(* IEC 61131-3 sources: plc-vscode/tests/st/test-ready/rusty/tests/lit/single/conversion, 6 files *)

(* ---- real_trunc_int.st ---- *)
// RUN: (%COMPILE %s && %RUN) | %CHECK %s
FUNCTION main
    printf('%d$N', REAL_TRUNC_SINT(5.6));       // CHECK: 5
    printf('%d$N', REAL_TRUNC_USINT(5.6));      // CHECK: 5
    printf('%d$N', REAL_TRUNC_INT(5.6));        // CHECK: 5
    printf('%d$N', REAL_TRUNC_UINT(5.6));       // CHECK: 5
    printf('%d$N', REAL_TRUNC_INT(5.6));        // CHECK: 5
    printf('%d$N', REAL_TRUNC_UINT(5.6));       // CHECK: 5
    printf('%d$N', REAL_TRUNC_DINT(5.6));       // CHECK: 5
    printf('%d$N', REAL_TRUNC_UDINT(5.6));      // CHECK: 5
    printf('%d$N', REAL_TRUNC_LINT(5.6));       // CHECK: 5
    printf('%d$N', REAL_TRUNC_ULINT(5.6));      // CHECK: 5

    printf('%d$N', REAL_TRUNC_SINT(-5.6));      // CHECK: -5
    printf('%d$N', REAL_TRUNC_INT(-5.6));       // CHECK: -5
    printf('%d$N', REAL_TRUNC_DINT(-5.6));      // CHECK: -5
    printf('%d$N', REAL_TRUNC_LINT(-5.6));      // CHECK: -5
END_FUNCTION

(* ---- to_bit.st ---- *)
// Note: Tests are kept simple because there are already tests covering the underliny X_TO_Y functions, which
//       the TO_Y(X) functions are based on.

// RUN: (%COMPILE %s && %RUN) | %CHECK %s
FUNCTION main
    printf('%d$N', TO_BOOL(BOOL#FALSE));        // CHECK: 0
    printf('%d$N', TO_BOOL(BOOL#TRUE));         // CHECK: 1
    printf('%d$N', TO_BOOL(BYTE#0));            // CHECK: 0
    printf('%d$N', TO_BOOL(BYTE#5));            // CHECK: 1
    printf('%d$N', TO_BOOL(WORD#0));            // CHECK: 0
    printf('%d$N', TO_BOOL(WORD#5));            // CHECK: 1
    printf('%d$N', TO_BOOL(DWORD#0));           // CHECK: 0
    printf('%d$N', TO_BOOL(DWORD#5));           // CHECK: 1
    printf('%d$N', TO_BOOL(LWORD#0));           // CHECK: 0
    printf('%d$N', TO_BOOL(LWORD#5));           // CHECK: 1

    printf('%d$N', TO_BYTE(BYTE#5));            // CHECK: 5
    printf('%d$N', TO_BYTE(BOOL#FALSE));        // CHECK: 0
    printf('%d$N', TO_BYTE(BOOL#TRUE));         // CHECK: 1
    printf('%d$N', TO_BYTE(CHAR#'a'));          // CHECK: 97
    printf('%d$N', TO_BYTE(WCHAR#"a"));         // CHECK: 97
    printf('%d$N', TO_BYTE(WORD#5));            // CHECK: 5
    printf('%d$N', TO_BYTE(DWORD#5));           // CHECK: 5
    printf('%d$N', TO_BYTE(LWORD#5));           // CHECK: 5

    printf('%d$N', TO_WORD(WORD#5));            // CHECK: 5
    printf('%d$N', TO_WORD(BOOL#FALSE));        // CHECK: 0
    printf('%d$N', TO_WORD(BOOL#TRUE));         // CHECK: 1
    printf('%d$N', TO_WORD(CHAR#'a'));          // CHECK: 97
    printf('%d$N', TO_WORD(WCHAR#"a"));         // CHECK: 97
    printf('%d$N', TO_WORD(BYTE#5));            // CHECK: 5
    printf('%d$N', TO_WORD(DWORD#5));           // CHECK: 5
    printf('%d$N', TO_WORD(LWORD#5));           // CHECK: 5

    printf('%d$N', TO_DWORD(DWORD#5));          // CHECK: 5
    printf('%d$N', TO_DWORD(BOOL#FALSE));       // CHECK: 0
    printf('%d$N', TO_DWORD(BOOL#TRUE));        // CHECK: 1
    printf('%d$N', TO_DWORD(CHAR#'a'));         // CHECK: 97
    printf('%d$N', TO_DWORD(WCHAR#'a'));        // CHECK: 97
    printf('%d$N', TO_DWORD(BYTE#5));           // CHECK: 5
    printf('%d$N', TO_DWORD(WORD#5));           // CHECK: 5
    printf('%d$N', TO_DWORD(LWORD#5));          // CHECK: 5

    printf('%d$N', TO_LWORD(LWORD#5));          // CHECK: 5
    printf('%d$N', TO_LWORD(BOOL#FALSE));       // CHECK: 0
    printf('%d$N', TO_LWORD(BOOL#TRUE));        // CHECK: 1
    printf('%d$N', TO_LWORD(CHAR#'a'));         // CHECK: 97
    printf('%d$N', TO_LWORD(WCHAR#'a'));        // CHECK: 97
    printf('%d$N', TO_LWORD(BYTE#5));           // CHECK: 5
    printf('%d$N', TO_LWORD(WORD#5));           // CHECK: 5
    printf('%d$N', TO_LWORD(DWORD#5));          // CHECK: 5
END_FUNCTION

(* ---- to_date_time.st ---- *)
// RUN: (%COMPILE %s && %RUN) | %CHECK %s
FUNCTION main
    // TO_TIME
    printf('%s$N', REF(TIME_TO_STRING(TO_TIME(LTIME#10s))));                        // CHECK: 10s

    // TO_LTIME
    printf('%s$N', REF(TIME_TO_STRING(TO_LTIME(TIME#10s))));                        // CHECK: 10s

    // TO_DT
    printf('%s$N', REF(TIME_TO_STRING(TO_DT(LDT#2024-11-12-16:36:15.100))));        // CHECK: 20039d16h36m15s100ms

    // TO_LDT
    printf('%s$N', REF(TIME_TO_STRING(TO_LDT(DT#2024-11-12-16:36:15.100))));        // CHECK: 20039d16h36m15s100ms

    // TO_DATE
    printf('%s$N', REF(TIME_TO_STRING(TO_DATE(DT#2024-11-12-16:36:15.100))));       // CHECK: 20039d
    printf('%s$N', REF(TIME_TO_STRING(TO_DATE(LDT#2024-11-12-16:36:15.100))));      // CHECK: 20039d

    // TO_LDATE
    printf('%s$N', REF(TIME_TO_STRING(TO_LDATE(DT#2024-11-12-16:36:15.100))));       // CHECK: 20039d
    printf('%s$N', REF(TIME_TO_STRING(TO_LDATE(LDT#2024-11-12-16:36:15.100))));      // CHECK: 20039d

    // TO_TOD
    printf('%s$N', REF(LTOD_TO_STRING(TO_TOD(LTOD#16:36:15))));                     // CHECK: 16:36:15
    printf('%s$N', REF(TOD_TO_STRING(TO_TOD(DT#2024-11-12-16:36:15.100))));         // CHECK: 16:36:15.100
    printf('%s$N', REF(TOD_TO_STRING(TO_TOD(LDT#2024-11-12-16:36:15.100))));        // CHECK: 16:36:15.100

    // TO_LTOD
    printf('%s$N', REF(LTOD_TO_STRING(TO_LTOD(TOD#16:36:15))));                     // CHECK: 16:36:15
    printf('%s$N', REF(LTOD_TO_STRING(TO_LTOD(DT#2024-11-12-16:36:15.100))));       // CHECK: 16:36:15.100
    printf('%s$N', REF(LTOD_TO_STRING(TO_LTOD(LDT#2024-11-12-16:36:15.100))));      // CHECK: 16:36:15.100
END_FUNCTION

(* ---- to_num.st ---- *)
// RUN: (%COMPILE %s && %RUN) | %CHECK %s
FUNCTION main
    printf('%d$N', TO_SINT(SINT#5));            // CHECK: 5
    printf('%d$N', TO_SINT(USINT#5));           // CHECK: 5
    printf('%d$N', TO_SINT(INT#5));             // CHECK: 5
    printf('%d$N', TO_SINT(UINT#5));            // CHECK: 5
    printf('%d$N', TO_SINT(DINT#5));            // CHECK: 5
    printf('%d$N', TO_SINT(UDINT#5));           // CHECK: 5
    printf('%d$N', TO_SINT(LINT#5));            // CHECK: 5
    printf('%d$N', TO_SINT(ULINT#5));           // CHECK: 5

    printf('%d$N', TO_USINT(SINT#5));            // CHECK: 5
    printf('%d$N', TO_USINT(USINT#5));           // CHECK: 5
    printf('%d$N', TO_USINT(INT#5));             // CHECK: 5
    printf('%d$N', TO_USINT(UINT#5));            // CHECK: 5
    printf('%d$N', TO_USINT(DINT#5));            // CHECK: 5
    printf('%d$N', TO_USINT(UDINT#5));           // CHECK: 5
    printf('%d$N', TO_USINT(LINT#5));            // CHECK: 5
    printf('%d$N', TO_USINT(ULINT#5));           // CHECK: 5

    printf('%d$N', TO_INT(SINT#5));            // CHECK: 5
    printf('%d$N', TO_INT(USINT#5));           // CHECK: 5
    printf('%d$N', TO_INT(INT#5));             // CHECK: 5
    printf('%d$N', TO_INT(UINT#5));            // CHECK: 5
    printf('%d$N', TO_INT(DINT#5));            // CHECK: 5
    printf('%d$N', TO_INT(UDINT#5));           // CHECK: 5
    printf('%d$N', TO_INT(LINT#5));            // CHECK: 5
    printf('%d$N', TO_INT(ULINT#5));           // CHECK: 5

    printf('%d$N', TO_UINT(SINT#5));            // CHECK: 5
    printf('%d$N', TO_UINT(USINT#5));           // CHECK: 5
    printf('%d$N', TO_UINT(INT#5));             // CHECK: 5
    printf('%d$N', TO_UINT(UINT#5));            // CHECK: 5
    printf('%d$N', TO_UINT(DINT#5));            // CHECK: 5
    printf('%d$N', TO_UINT(UDINT#5));           // CHECK: 5
    printf('%d$N', TO_UINT(LINT#5));            // CHECK: 5
    printf('%d$N', TO_UINT(ULINT#5));           // CHECK: 5

    printf('%d$N', TO_DINT(SINT#5));            // CHECK: 5
    printf('%d$N', TO_DINT(USINT#5));           // CHECK: 5
    printf('%d$N', TO_DINT(INT#5));             // CHECK: 5
    printf('%d$N', TO_DINT(UINT#5));            // CHECK: 5
    printf('%d$N', TO_DINT(DINT#5));            // CHECK: 5
    printf('%d$N', TO_DINT(UDINT#5));           // CHECK: 5
    printf('%d$N', TO_DINT(LINT#5));            // CHECK: 5
    printf('%d$N', TO_DINT(ULINT#5));           // CHECK: 5

    printf('%d$N', TO_UDINT(SINT#5));            // CHECK: 5
    printf('%d$N', TO_UDINT(USINT#5));           // CHECK: 5
    printf('%d$N', TO_UDINT(INT#5));             // CHECK: 5
    printf('%d$N', TO_UDINT(UINT#5));            // CHECK: 5
    printf('%d$N', TO_UDINT(DINT#5));            // CHECK: 5
    printf('%d$N', TO_UDINT(UDINT#5));           // CHECK: 5
    printf('%d$N', TO_UDINT(LINT#5));            // CHECK: 5
    printf('%d$N', TO_UDINT(ULINT#5));           // CHECK: 5

    printf('%d$N', TO_LINT(SINT#5));            // CHECK: 5
    printf('%d$N', TO_LINT(USINT#5));           // CHECK: 5
    printf('%d$N', TO_LINT(INT#5));             // CHECK: 5
    printf('%d$N', TO_LINT(UINT#5));            // CHECK: 5
    printf('%d$N', TO_LINT(DINT#5));            // CHECK: 5
    printf('%d$N', TO_LINT(UDINT#5));           // CHECK: 5
    printf('%d$N', TO_LINT(LINT#5));            // CHECK: 5
    printf('%d$N', TO_LINT(ULINT#5));           // CHECK: 5

    printf('%d$N', TO_ULINT(SINT#5));            // CHECK: 5
    printf('%d$N', TO_ULINT(USINT#5));           // CHECK: 5
    printf('%d$N', TO_ULINT(INT#5));             // CHECK: 5
    printf('%d$N', TO_ULINT(UINT#5));            // CHECK: 5
    printf('%d$N', TO_ULINT(DINT#5));            // CHECK: 5
    printf('%d$N', TO_ULINT(UDINT#5));           // CHECK: 5
    printf('%d$N', TO_ULINT(LINT#5));            // CHECK: 5
    printf('%d$N', TO_ULINT(ULINT#5));           // CHECK: 5

    // REAL and LREAL tests, where we want to see rounding

    printf('%d$N', TO_SINT(REAL#4.0));          // CHECK: 4
    printf('%d$N', TO_SINT(REAL#4.1));          // CHECK: 4
    printf('%d$N', TO_SINT(REAL#4.2));          // CHECK: 4
    printf('%d$N', TO_SINT(REAL#4.3));          // CHECK: 4
    printf('%d$N', TO_SINT(REAL#4.4));          // CHECK: 4
    printf('%d$N', TO_SINT(REAL#4.5));          // CHECK: 5
    printf('%d$N', TO_SINT(REAL#4.6));          // CHECK: 5
    printf('%d$N', TO_SINT(REAL#4.7));          // CHECK: 5
    printf('%d$N', TO_SINT(REAL#4.8));          // CHECK: 5
    printf('%d$N', TO_SINT(REAL#4.9));          // CHECK: 5
    printf('%d$N', TO_SINT(LREAL#4.0));         // CHECK: 4
    printf('%d$N', TO_SINT(LREAL#4.1));         // CHECK: 4
    printf('%d$N', TO_SINT(LREAL#4.2));         // CHECK: 4
    printf('%d$N', TO_SINT(LREAL#4.3));         // CHECK: 4
    printf('%d$N', TO_SINT(LREAL#4.4));         // CHECK: 4
    printf('%d$N', TO_SINT(LREAL#4.5));         // CHECK: 5
    printf('%d$N', TO_SINT(LREAL#4.6));         // CHECK: 5
    printf('%d$N', TO_SINT(LREAL#4.7));         // CHECK: 5
    printf('%d$N', TO_SINT(LREAL#4.8));         // CHECK: 5
    printf('%d$N', TO_SINT(LREAL#4.9));         // CHECK: 5

    printf('%d$N', TO_USINT(REAL#4.0));          // CHECK: 4
    printf('%d$N', TO_USINT(REAL#4.1));          // CHECK: 4
    printf('%d$N', TO_USINT(REAL#4.2));          // CHECK: 4
    printf('%d$N', TO_USINT(REAL#4.3));          // CHECK: 4
    printf('%d$N', TO_USINT(REAL#4.4));          // CHECK: 4
    printf('%d$N', TO_USINT(REAL#4.5));          // CHECK: 5
    printf('%d$N', TO_USINT(REAL#4.6));          // CHECK: 5
    printf('%d$N', TO_USINT(REAL#4.7));          // CHECK: 5
    printf('%d$N', TO_USINT(REAL#4.8));          // CHECK: 5
    printf('%d$N', TO_USINT(REAL#4.9));          // CHECK: 5
    printf('%d$N', TO_USINT(LREAL#4.0));         // CHECK: 4
    printf('%d$N', TO_USINT(LREAL#4.1));         // CHECK: 4
    printf('%d$N', TO_USINT(LREAL#4.2));         // CHECK: 4
    printf('%d$N', TO_USINT(LREAL#4.3));         // CHECK: 4
    printf('%d$N', TO_USINT(LREAL#4.4));         // CHECK: 4
    printf('%d$N', TO_USINT(LREAL#4.5));         // CHECK: 5
    printf('%d$N', TO_USINT(LREAL#4.6));         // CHECK: 5
    printf('%d$N', TO_USINT(LREAL#4.7));         // CHECK: 5
    printf('%d$N', TO_USINT(LREAL#4.8));         // CHECK: 5
    printf('%d$N', TO_USINT(LREAL#4.9));         // CHECK: 5

    printf('%d$N', TO_INT(REAL#4.0));          // CHECK: 4
    printf('%d$N', TO_INT(REAL#4.1));          // CHECK: 4
    printf('%d$N', TO_INT(REAL#4.2));          // CHECK: 4
    printf('%d$N', TO_INT(REAL#4.3));          // CHECK: 4
    printf('%d$N', TO_INT(REAL#4.4));          // CHECK: 4
    printf('%d$N', TO_INT(REAL#4.5));          // CHECK: 5
    printf('%d$N', TO_INT(REAL#4.6));          // CHECK: 5
    printf('%d$N', TO_INT(REAL#4.7));          // CHECK: 5
    printf('%d$N', TO_INT(REAL#4.8));          // CHECK: 5
    printf('%d$N', TO_INT(REAL#4.9));          // CHECK: 5
    printf('%d$N', TO_INT(LREAL#4.0));         // CHECK: 4
    printf('%d$N', TO_INT(LREAL#4.1));         // CHECK: 4
    printf('%d$N', TO_INT(LREAL#4.2));         // CHECK: 4
    printf('%d$N', TO_INT(LREAL#4.3));         // CHECK: 4
    printf('%d$N', TO_INT(LREAL#4.4));         // CHECK: 4
    printf('%d$N', TO_INT(LREAL#4.5));         // CHECK: 5
    printf('%d$N', TO_INT(LREAL#4.6));         // CHECK: 5
    printf('%d$N', TO_INT(LREAL#4.7));         // CHECK: 5
    printf('%d$N', TO_INT(LREAL#4.8));         // CHECK: 5
    printf('%d$N', TO_INT(LREAL#4.9));         // CHECK: 5

    printf('%d$N', TO_UINT(REAL#4.0));          // CHECK: 4
    printf('%d$N', TO_UINT(REAL#4.1));          // CHECK: 4
    printf('%d$N', TO_UINT(REAL#4.2));          // CHECK: 4
    printf('%d$N', TO_UINT(REAL#4.3));          // CHECK: 4
    printf('%d$N', TO_UINT(REAL#4.4));          // CHECK: 4
    printf('%d$N', TO_UINT(REAL#4.5));          // CHECK: 5
    printf('%d$N', TO_UINT(REAL#4.6));          // CHECK: 5
    printf('%d$N', TO_UINT(REAL#4.7));          // CHECK: 5
    printf('%d$N', TO_UINT(REAL#4.8));          // CHECK: 5
    printf('%d$N', TO_UINT(REAL#4.9));          // CHECK: 5
    printf('%d$N', TO_UINT(LREAL#4.0));         // CHECK: 4
    printf('%d$N', TO_UINT(LREAL#4.1));         // CHECK: 4
    printf('%d$N', TO_UINT(LREAL#4.2));         // CHECK: 4
    printf('%d$N', TO_UINT(LREAL#4.3));         // CHECK: 4
    printf('%d$N', TO_UINT(LREAL#4.4));         // CHECK: 4
    printf('%d$N', TO_UINT(LREAL#4.5));         // CHECK: 5
    printf('%d$N', TO_UINT(LREAL#4.6));         // CHECK: 5
    printf('%d$N', TO_UINT(LREAL#4.7));         // CHECK: 5
    printf('%d$N', TO_UINT(LREAL#4.8));         // CHECK: 5
    printf('%d$N', TO_UINT(LREAL#4.9));         // CHECK: 5

    printf('%d$N', TO_DINT(REAL#4.0));          // CHECK: 4
    printf('%d$N', TO_DINT(REAL#4.1));          // CHECK: 4
    printf('%d$N', TO_DINT(REAL#4.2));          // CHECK: 4
    printf('%d$N', TO_DINT(REAL#4.3));          // CHECK: 4
    printf('%d$N', TO_DINT(REAL#4.4));          // CHECK: 4
    printf('%d$N', TO_DINT(REAL#4.5));          // CHECK: 5
    printf('%d$N', TO_DINT(REAL#4.6));          // CHECK: 5
    printf('%d$N', TO_DINT(REAL#4.7));          // CHECK: 5
    printf('%d$N', TO_DINT(REAL#4.8));          // CHECK: 5
    printf('%d$N', TO_DINT(REAL#4.9));          // CHECK: 5
    printf('%d$N', TO_DINT(LREAL#4.0));         // CHECK: 4
    printf('%d$N', TO_DINT(LREAL#4.1));         // CHECK: 4
    printf('%d$N', TO_DINT(LREAL#4.2));         // CHECK: 4
    printf('%d$N', TO_DINT(LREAL#4.3));         // CHECK: 4
    printf('%d$N', TO_DINT(LREAL#4.4));         // CHECK: 4
    printf('%d$N', TO_DINT(LREAL#4.5));         // CHECK: 5
    printf('%d$N', TO_DINT(LREAL#4.6));         // CHECK: 5
    printf('%d$N', TO_DINT(LREAL#4.7));         // CHECK: 5
    printf('%d$N', TO_DINT(LREAL#4.8));         // CHECK: 5
    printf('%d$N', TO_DINT(LREAL#4.9));         // CHECK: 5

    printf('%d$N', TO_UDINT(REAL#4.0));          // CHECK: 4
    printf('%d$N', TO_UDINT(REAL#4.1));          // CHECK: 4
    printf('%d$N', TO_UDINT(REAL#4.2));          // CHECK: 4
    printf('%d$N', TO_UDINT(REAL#4.3));          // CHECK: 4
    printf('%d$N', TO_UDINT(REAL#4.4));          // CHECK: 4
    printf('%d$N', TO_UDINT(REAL#4.5));          // CHECK: 5
    printf('%d$N', TO_UDINT(REAL#4.6));          // CHECK: 5
    printf('%d$N', TO_UDINT(REAL#4.7));          // CHECK: 5
    printf('%d$N', TO_UDINT(REAL#4.8));          // CHECK: 5
    printf('%d$N', TO_UDINT(REAL#4.9));          // CHECK: 5
    printf('%d$N', TO_UDINT(LREAL#4.0));         // CHECK: 4
    printf('%d$N', TO_UDINT(LREAL#4.1));         // CHECK: 4
    printf('%d$N', TO_UDINT(LREAL#4.2));         // CHECK: 4
    printf('%d$N', TO_UDINT(LREAL#4.3));         // CHECK: 4
    printf('%d$N', TO_UDINT(LREAL#4.4));         // CHECK: 4
    printf('%d$N', TO_UDINT(LREAL#4.5));         // CHECK: 5
    printf('%d$N', TO_UDINT(LREAL#4.6));         // CHECK: 5
    printf('%d$N', TO_UDINT(LREAL#4.7));         // CHECK: 5
    printf('%d$N', TO_UDINT(LREAL#4.8));         // CHECK: 5
    printf('%d$N', TO_UDINT(LREAL#4.9));         // CHECK: 5

    printf('%d$N', TO_LINT(REAL#4.0));          // CHECK: 4
    printf('%d$N', TO_LINT(REAL#4.1));          // CHECK: 4
    printf('%d$N', TO_LINT(REAL#4.2));          // CHECK: 4
    printf('%d$N', TO_LINT(REAL#4.3));          // CHECK: 4
    printf('%d$N', TO_LINT(REAL#4.4));          // CHECK: 4
    printf('%d$N', TO_LINT(REAL#4.5));          // CHECK: 5
    printf('%d$N', TO_LINT(REAL#4.6));          // CHECK: 5
    printf('%d$N', TO_LINT(REAL#4.7));          // CHECK: 5
    printf('%d$N', TO_LINT(REAL#4.8));          // CHECK: 5
    printf('%d$N', TO_LINT(REAL#4.9));          // CHECK: 5
    printf('%d$N', TO_LINT(LREAL#4.0));         // CHECK: 4
    printf('%d$N', TO_LINT(LREAL#4.1));         // CHECK: 4
    printf('%d$N', TO_LINT(LREAL#4.2));         // CHECK: 4
    printf('%d$N', TO_LINT(LREAL#4.3));         // CHECK: 4
    printf('%d$N', TO_LINT(LREAL#4.4));         // CHECK: 4
    printf('%d$N', TO_LINT(LREAL#4.5));         // CHECK: 5
    printf('%d$N', TO_LINT(LREAL#4.6));         // CHECK: 5
    printf('%d$N', TO_LINT(LREAL#4.7));         // CHECK: 5
    printf('%d$N', TO_LINT(LREAL#4.8));         // CHECK: 5
    printf('%d$N', TO_LINT(LREAL#4.9));         // CHECK: 5

    printf('%d$N', TO_ULINT(REAL#4.0));          // CHECK: 4
    printf('%d$N', TO_ULINT(REAL#4.1));          // CHECK: 4
    printf('%d$N', TO_ULINT(REAL#4.2));          // CHECK: 4
    printf('%d$N', TO_ULINT(REAL#4.3));          // CHECK: 4
    printf('%d$N', TO_ULINT(REAL#4.4));          // CHECK: 4
    printf('%d$N', TO_ULINT(REAL#4.5));          // CHECK: 5
    printf('%d$N', TO_ULINT(REAL#4.6));          // CHECK: 5
    printf('%d$N', TO_ULINT(REAL#4.7));          // CHECK: 5
    printf('%d$N', TO_ULINT(REAL#4.8));          // CHECK: 5
    printf('%d$N', TO_ULINT(REAL#4.9));          // CHECK: 5
    printf('%d$N', TO_ULINT(LREAL#4.0));         // CHECK: 4
    printf('%d$N', TO_ULINT(LREAL#4.1));         // CHECK: 4
    printf('%d$N', TO_ULINT(LREAL#4.2));         // CHECK: 4
    printf('%d$N', TO_ULINT(LREAL#4.3));         // CHECK: 4
    printf('%d$N', TO_ULINT(LREAL#4.4));         // CHECK: 4
    printf('%d$N', TO_ULINT(LREAL#4.5));         // CHECK: 5
    printf('%d$N', TO_ULINT(LREAL#4.6));         // CHECK: 5
    printf('%d$N', TO_ULINT(LREAL#4.7));         // CHECK: 5
    printf('%d$N', TO_ULINT(LREAL#4.8));         // CHECK: 5
    printf('%d$N', TO_ULINT(LREAL#4.9));         // CHECK: 5
END_FUNCTION

(* ---- to_string.st ---- *)
// RUN: (%COMPILE %s && %RUN) | %CHECK %s
FUNCTION main : DINT
    // TO_CHAR
    printf('%c$N', TO_CHAR(WCHAR#"a"));             // CHECK: a
    printf('%c$N', TO_CHAR(STRING#'foo'));          // CHECK: f

    // TO_WCHAR
    printf('%c$N', TO_WCHAR(CHAR#'a'));             // CHECK: a
    printf('%c$N', TO_WCHAR(WSTRING#"foo"));        // CHECK: f

    // TO_STRING
    printf('%s$N', REF(TO_STRING(CHAR#'a')));       // CHECK: a
    printf('%s$N', REF(TO_STRING(WSTRING#"foo")));  // CHECK: foo

    // TO_WSTRING
    printf('%s$N', REF(TO_STRING(TO_WSTRING(WCHAR#"a"))));      // CHECK: a
    printf('%s$N', REF(TO_STRING(TO_WSTRING(STRING#'foo'))));   // CHECK: foo
END_FUNCTION

(* ---- trunc_int.st ---- *)
// RUN: (%COMPILE %s && %RUN) | %CHECK %s
FUNCTION main
    // REAL
    printf('%d$N', TRUNC_SINT(REAL#5.6));       // CHECK: 5
    printf('%d$N', TRUNC_USINT(REAL#5.6));      // CHECK: 5
    printf('%d$N', TRUNC_INT(REAL#5.6));        // CHECK: 5
    printf('%d$N', TRUNC_UINT(REAL#5.6));       // CHECK: 5
    printf('%d$N', TRUNC_INT(REAL#5.6));        // CHECK: 5
    printf('%d$N', TRUNC_UINT(REAL#5.6));       // CHECK: 5
    printf('%d$N', TRUNC_DINT(REAL#5.6));       // CHECK: 5
    printf('%d$N', TRUNC_UDINT(REAL#5.6));      // CHECK: 5
    printf('%d$N', TRUNC_LINT(REAL#5.6));       // CHECK: 5
    printf('%d$N', TRUNC_ULINT(REAL#5.6));      // CHECK: 5

    printf('%d$N', TRUNC_SINT(REAL#-5.6));      // CHECK: -5
    printf('%d$N', TRUNC_INT(REAL#-5.6));       // CHECK: -5
    printf('%d$N', TRUNC_DINT(REAL#-5.6));      // CHECK: -5
    printf('%d$N', TRUNC_LINT(REAL#-5.6));      // CHECK: -5

    // LREAL
    printf('%d$N', TRUNC_SINT(LREAL#5.6));       // CHECK: 5
    printf('%d$N', TRUNC_USINT(LREAL#5.6));      // CHECK: 5
    printf('%d$N', TRUNC_INT(LREAL#5.6));        // CHECK: 5
    printf('%d$N', TRUNC_UINT(LREAL#5.6));       // CHECK: 5
    printf('%d$N', TRUNC_INT(LREAL#5.6));        // CHECK: 5
    printf('%d$N', TRUNC_UINT(LREAL#5.6));       // CHECK: 5
    printf('%d$N', TRUNC_DINT(LREAL#5.6));       // CHECK: 5
    printf('%d$N', TRUNC_UDINT(LREAL#5.6));      // CHECK: 5
    printf('%d$N', TRUNC_LINT(LREAL#5.6));       // CHECK: 5
    printf('%d$N', TRUNC_ULINT(LREAL#5.6));      // CHECK: 5

    printf('%d$N', TRUNC_SINT(LREAL#-5.6));      // CHECK: -5
    printf('%d$N', TRUNC_INT(LREAL#-5.6));       // CHECK: -5
    printf('%d$N', TRUNC_DINT(LREAL#-5.6));      // CHECK: -5
    printf('%d$N', TRUNC_LINT(LREAL#-5.6));      // CHECK: -5
END_FUNCTION
